{region 'Documentation'}
(*!
<summary>Checks equality with the expected WORD value.</summary>
*)
{endregion}
FUNCTION_BLOCK AssertEqual_Word EXTENDS AssertionBase
VAR_INPUT
    IN : WORD; //! Actual value checked or observed by this Assertion.
    Expected : WORD; //! Reference value for comparison with IN.
END_VAR

SUPER^();

{region 'Documentation'}
(*!
<summary>Check equality with the expected WORD value.</summary>
*)
{endregion}
METHOD PROTECTED Assert
VAR
    Message : STRING(GVL_Constants.MessageLength);
    ExpectedText : STRING(GVL_Constants.AssertionValueLength);
    ActualText : STRING(GVL_Constants.AssertionValueLength);
END_VAR
VAR CONSTANT
    HexDigitCount : USINT := 4;
END_VAR
IF NOT EvaluationActive THEN
    RETURN;
END_IF;

IF Result = E_Result.Error THEN
    RETURN;
END_IF;

IF Result = E_Result.Failed THEN
    RETURN;
END_IF;

IF IN <> Expected THEN
    ExpectedText := CreateAssertionTextValue_Hex(Value := WORD_TO_LWORD(Expected),
        DigitCount := HexDigitCount);
    ActualText := CreateAssertionTextValue_Hex(Value := WORD_TO_LWORD(IN),
        DigitCount := HexDigitCount);
    Message := CONCAT('Assertion failed: values are not equal. Expected = ',
        ExpectedText);
    Message := CONCAT(Message, ', Actual = ');
    Message := CONCAT(Message, ActualText);
    Message := CONCAT(Message, '.');
    Fail(Message := Message);
    RETURN;
END_IF;

Pass();
END_METHOD

END_FUNCTION_BLOCK

(* stored: Version 1.1.0.1
   POU AssertEqual_Word: Id {42fe4084-717d-450b-b595-9762fa2c3b97}, SpecialFunc None
   Folder Internal: Id {86262986-83f4-4fa9-9517-7a7de02f976d}
   Method Assert: Id {c7757eab-e7a0-4811-ac58-ae226e427148} *)
